TYPE "ST_PressDemoOutImm"
VERSION : 0.1
   STRUCT
      Homed : Bool;
   END_STRUCT;

END_TYPE

